Fanuc KAREL source: ko00062.KL

-- PROVISIONAL review KL for V770-1; original PC SHA256 d1c0714e1dde4b1aef707c0355f217c5fd76b1a177c6e8051ada0fe2c039fbf9
-- Incomplete behavior may be omitted. Consult companion uncertainty JSON. Do not deploy.
PROGRAM KO00062
%NOLOCKGROUP
BEGIN
  -- UNRESOLVED_PC offsets 5-12; opcodes 9D,23
  -- UNRESOLVED_PC offsets 17-69; opcodes 27,27,49,7E,AD,27,49,7E,AD,22,31,7E,4A
  -- UNRESOLVED_PC offsets 74-78; opcodes 7F
END KO00062
